{attribute 'qualified_only'}
VAR_GLOBAL RETAIN
	LightH1Config : stLightConfig := (
		BrightnessSmoothTime := T#2S);
END_VAR

(* stored: Version 1.1.0.1
   GVL gvlLights: Id {dd61c03b-2734-4b8a-940c-ae1964cdd439} *)
